(* IEC 61131-3 sources: generating_plc_code_with_llms/Code#1/Platypus2/third run, 5 files *)

(* ---- 12.st ---- *)
// 9.175787448883057s
// 1
function sinh(x)
    return exp(x)*cosh(x);
end_function

(* ---- 13.st ---- *)
// 20.42183232307434s
// 2
REPEAT
    IF (SELECTED_NUMBER = 10) THEN
        EXIT
    END_IF
END_REPEAT

(* ---- 15.st ---- *)
// 32.1113395690918s
// 2
IF (E_A = 0) THEN
    IF (P_HU = 0 AND P_AL = 1) THEN
        P_AL = 0
    END_IF
END_IF

(* ---- 17.st ---- *)
// 79.89235615730286s
// 2
IF (HUMIDITY < 40 OR HUMIDITY > 75) THEN
    DISPLAY "Humidity out of range!"
ELSEIF (TEMPERATURE < 18 OR TEMPERATURE > 25) THEN
    IF (TEMPERATURE < 18) THEN
        DISPLAY "Cold"
    ELSEIF (TEMPERATURE > 25) THEN
        DISPLAY "Hot"
    END_IF
ELSE
    IF (HUMIDITY BETWEEN 40 AND 75 AND TEMPERATURE BETWEEN 18 AND 25) THEN
        DISPLAY "Opt"
    ELSE
        DISPLAY "Temp. OK"
    END_IF
END_IF

(* ---- 19.st ---- *)
// 69.78339076042175s
// 2
```
THICKNESS(MD_1)
D_MAX := MD_1;
D_MIN := MD_1;
IF (S1 = 0) THEN
    IF (D_MAX > V_MAX OR D_MIN < V_MIN) THEN
        P1 := TRUE;
    ELSE
        P1 := FALSE;
    END_IF;
END_IF;
```
